(* IEC 61131-3 sources: plc-st-coding-agent/progress/evidence/f14_p1_20261111b/jobs/custom_minimax-m27 (part 2) *)

(* ---- self-hard-06.candidate_01.st ---- *)
FUNCTION_BLOCK FB
VAR_INPUT
    runRequest        : BOOL;
    pressure          : REAL;
    pressureValid     : BOOL;
    fuelFlow          : REAL;
    steamFlow         : REAL;
    outletCmd         : INT;
    outletFeedback    : INT;
    resetBtn          : BOOL;
END_VAR
VAR_OUTPUT
    tripLatched       : BOOL;
    fuelPermit        : BOOL;
    currentCauseMask  : WORD;
    latchedCauseMask  : WORD;
    diagnosticActive  : BOOL;
END_VAR
VAR
    stuckCount   : INT  := 0;      (* consecutive cycles for valve‑stuck detection *)
    prevResetBtn : BOOL := FALSE;   (* previous state of reset button *)
END_VAR

(* ------------------------------------------------------------------
   1. Valve‑stuck consecutive‑cycle detection
   ------------------------------------------------------------------ *)
IF runRequest AND pressureValid AND (pressure >= 4500.0)
   AND (outletCmd >= 50) AND (outletFeedback <= 10) THEN
    IF stuckCount < 3 THEN
        stuckCount := stuckCount + 1;
    END_IF;
ELSE
    stuckCount := 0;
END_IF;

(* ------------------------------------------------------------------
   2. Current cause mask (bits 0…3)
   ------------------------------------------------------------------ *)
IF NOT runRequest THEN
    currentCauseMask := 0;                     (* S5 *)

ELSIF NOT pressureValid THEN
    currentCauseMask := 1;                     (* bit0 – transmitter failure, S12 *)

ELSE
    (* pressureValid = TRUE *)
    IF pressure >= 4500.0 THEN
        (* Over‑pressure – evaluate bit1 (valve stuck) and bit2 (combustion excess) *)
        currentCauseMask := 0;

        IF stuckCount >= 3 THEN
            currentCauseMask := 2;             (* bit1 *)
        END_IF;

        IF (fuelFlow >= 4.0) AND (steamFlow <= 10.0) THEN
            currentCauseMask := currentCauseMask OR 4;  (* bit2 *)
        END_IF;

        (* If neither cause is identified, set bit3 (unlocated) *)
        IF currentCauseMask = 0 THEN
            currentCauseMask := 8;             (* bit3 *)
        END_IF;
    ELSE
        currentCauseMask := 0;                 (* S6 *)
    END_IF;
END_IF;

(* ------------------------------------------------------------------
   3. Trip condition
   ------------------------------------------------------------------ *)
(*  runRequest  AND ( pressureValid = FALSE  OR  pressure >= 4500.0 ) *)
tripLatched := tripLatched OR (runRequest AND (NOT pressureValid OR (pressure >= 4500.0)));

(* ------------------------------------------------------------------
   4. Reset on rising edge of reset button when conditions are met
   ------------------------------------------------------------------ *)
IF resetBtn AND NOT prevResetBtn AND NOT runRequest AND pressureValid AND (pressure <= 4200.0) THEN
    tripLatched := FALSE;
END_IF;
prevResetBtn := resetBtn;

(* ------------------------------------------------------------------
   5. Fuel permit
   ------------------------------------------------------------------ *)
fuelPermit := runRequest AND NOT tripLatched;   (* S3, N10‑S16 *)

(* ------------------------------------------------------------------
   6. Diagnostic active flag
   ------------------------------------------------------------------ *)
diagnosticActive := (currentCauseMask <> 0);    (* S7 *)

(* ------------------------------------------------------------------
   7. Accumulate cause mask while trip is latched
   ------------------------------------------------------------------ *)
IF tripLatched THEN
    latchedCauseMask := latchedCauseMask OR currentCauseMask;
ELSE
    latchedCauseMask := 0;                      (* N10‑S18 *)
END_IF;

END_FUNCTION_BLOCK

(* ---- self-medium-01.candidate_01.st ---- *)
TYPE ST_Recipe :
STRUCT
    recipeID   : INT;
    totalRatio : REAL;
    temperature: REAL;
END_STRUCT
END_TYPE

FUNCTION_BLOCK FB
VAR_INPUT
    recipe   : ARRAY[1..8] OF ST_Recipe;
    selSlot  : INT;
    loadCmd  : BOOL;
    running  : BOOL;
END_VAR
VAR_OUTPUT
    valid    : BOOL;
    loadedID : INT;
END_VAR
VAR
    prevLoadCmd  : BOOL := FALSE;
    prevRunning  : BOOL := FALSE;
    prevLoadedID : INT  := 0;
    prevValid    : BOOL := FALSE;
END_VAR
VAR_TEMP
    risingLoadCmd : BOOL;
    tmpRecipe     : ST_Recipe;
END_VAR

    // 检测 loadCmd 上升沿
    risingLoadCmd := loadCmd AND NOT prevLoadCmd;

    // 装载逻辑
    IF NOT running AND risingLoadCmd THEN
        // 槽位越界检查：必须先检查，不得访问数组外内存
        IF selSlot < 1 OR selSlot > 8 THEN
            valid   := FALSE;
            loadedID := 0;
        ELSE
            tmpRecipe := recipe[selSlot];
            // 槽位为空检查
            IF tmpRecipe.recipeID = 0 THEN
                valid   := FALSE;
                loadedID := 0;
            // 总配比越界检查 (99.0 <= totalRatio <= 101.0)
            ELSIF tmpRecipe.totalRatio < 99.0 OR tmpRecipe.totalRatio > 101.0 THEN
                valid   := FALSE;
                loadedID := 0;
            // 温度越界检查 (30.0 <= temperature <= 180.0)
            ELSIF tmpRecipe.temperature < 30.0 OR tmpRecipe.temperature > 180.0 THEN
                valid   := FALSE;
                loadedID := 0;
            ELSE
                valid    := TRUE;
                loadedID := tmpRecipe.recipeID;
            END_IF
        END_IF
    ELSE
        // 非装载周期：保持上一拍的值 (包括 running 状态)
        valid    := prevValid;
        loadedID := prevLoadedID;
    END_IF

    // 更新历史状态
    prevLoadCmd  := loadCmd;
    prevRunning  := running;
    prevLoadedID := loadedID;
    prevValid    := valid;

END_FUNCTION_BLOCK

(* ---- self-medium-02.candidate_01.st ---- *)
FUNCTION_BLOCK FB
VAR_INPUT
    enable    : BOOL;      (* 滤波使能，FALSE 时清空历史 *)
    rawValue  : REAL;      (* 本周期原始采样值 *)
END_VAR

VAR_OUTPUT
    filteredValue : REAL;  (* 滤波输出 *)
    windowFull    : BOOL;  (* 历史窗口已填满 8 个样本后置 TRUE *)
    sampleCount   : INT;   (* 当前窗口内有效样本数 0..8 *)
END_VAR

VAR
    buffer : ARRAY[0..7] OF REAL;  (* 8 点环形缓冲区 *)
    head   : INT := 0;             (* 下一写入位置 0..7 *)
    count  : INT := 0;             (* 有效样本数 0..8 *)
    full   : BOOL := FALSE;        (* 内部满窗标志 *)
END_VAR

VAR_TEMP
    sum : REAL;                    (* 临时累加和 *)
    idx : INT;                     (* 遍历索引 *)
    i   : INT;                     (* 循环计数器 *)
END_VAR

(*--------------------------------------------------------------------*)
(* 功能块主体                                                         *)
(*--------------------------------------------------------------------*)
IF enable THEN
    (* ----- 把新样本压入环形缓冲区 ----- *)
    buffer[head] := rawValue;                 (* 写入 *)
    head := (head + 1) MOD 8;                (* 头指针前移 *)
    IF count < 8 THEN
        count := count + 1;                  (* 样本计数 +1 *)
    END_IF
    full := (count = 8);                     (* 满窗标志 *)

ELSE
    (* ----- enable = FALSE：立即清零计数与满窗标志 ----- *)
    count := 0;
    full  := FALSE;
    (* head 保持不变，下一次 enable=TRUE 时会被覆盖 *)
END_IF

(* ----- 计算滤波输出（仅在有有效样本时） ----- *)
IF enable AND count > 0 THEN
    sum := 0.0;
    (*  oldest  = head - count (模 8) *)
    idx := (head - count + 8) MOD 8;
    FOR i := 0 TO count - 1 DO
        sum := sum + buffer[idx];
        idx := (idx + 1) MOD 8;
    END_FOR
    filteredValue := sum / INT_TO_REAL(count);   (* 算术平均 *)
END_IF
(* 当 enable=FALSE 时 filteredValue 保持不变 *)

(* ----- 输出信号 ----- *)
windowFull  := full;
sampleCount := count;

END_FUNCTION_BLOCK

(* ---- self-medium-03.candidate_01.st ---- *)
FUNCTION_BLOCK FB
VAR_INPUT
    openBtn    : BOOL;
    closeBtn   : BOOL;
    openLimit  : BOOL;
    closeLimit : BOOL;
    obstacle   : BOOL;
END_VAR

VAR_OUTPUT
    motorUp    : BOOL;
    motorDown  : BOOL;
    errorFlag  : BOOL;
END_VAR

VAR
    openBtnPrev    : BOOL := FALSE;
    closeBtnPrev   : BOOL := FALSE;
    combinedPrev   : BOOL := FALSE;
    prevMotorUp    : BOOL := FALSE;
    prevMotorDown  : BOOL := FALSE;
    prevErrorFlag  : BOOL := FALSE;
    state          : INT  := 0;   // 0=IDLE,1=OPENING,2=CLOSING,3=FAULT
END_VAR

(* Local auxiliary variables *)
VAR
    risingOpen     : BOOL;
    risingClose    : BOOL;
    risingCombined : BOOL;
    combinedNow    : BOOL;
    startOpen      : BOOL;
    startClose     : BOOL;
END_VAR

(* Detect combined button state *)
combinedNow    := openBtn AND closeBtn;

(* Detect rising edges *)
risingOpen     := openBtn   AND NOT openBtnPrev;
risingClose    := closeBtn  AND NOT closeBtnPrev;
risingCombined := combinedNow AND NOT combinedPrev;

(* Start conditions: new command from IDLE without fault and no obstacle *)
startOpen  := NOT prevMotorUp   AND NOT prevMotorDown   AND NOT prevErrorFlag
              AND risingOpen    AND NOT closeBtn AND NOT openLimit;

startClose := NOT prevMotorUp   AND NOT prevMotorDown   AND NOT prevErrorFlag
              AND risingClose   AND NOT openBtn  AND NOT closeLimit;

(* Motor commands according to S12 / S13 *)
motorUp   := NOT obstacle AND NOT openLimit
             AND (prevMotorUp OR startOpen);

motorDown := NOT obstacle AND NOT closeLimit
             AND (prevMotorDown OR startClose);

(* Error flag latch (S14) *)
errorFlag := obstacle OR (prevErrorFlag AND NOT risingCombined);

(* Optional state for external monitoring *)
IF errorFlag THEN
    state := 3;               (* FAULT *)
ELSIF motorUp THEN
    state := 1;               (* OPENING *)
ELSIF motorDown THEN
    state := 2;               (* CLOSING *)
ELSE
    state := 0;               (* IDLE *)
END_IF

(* Update previous values for next scan *)
openBtnPrev    := openBtn;
closeBtnPrev   := closeBtn;
combinedPrev   := combinedNow;
prevMotorUp    := motorUp;
prevMotorDown  := motorDown;
prevErrorFlag  := errorFlag;

END_FUNCTION_BLOCK

(* ---- self-medium-04.candidate_01.st ---- *)
FUNCTION_BLOCK FB
VAR_INPUT
    startBtn   : BOOL;
    resetBtn   : BOOL;
    doneSensor : BOOL;
    targetVol  : REAL;
    flowVol    : REAL;
END_VAR
VAR_OUTPUT
    valveOpen  : BOOL;
    fillsToday : INT;
END_VAR
VAR
    prev_startBtn   : BOOL := FALSE;
    prev_resetBtn   : BOOL := FALSE;
    prev_valveOpen  : BOOL := FALSE;
    currentFillVol  : REAL := 0.0;
    pendingConfirm  : BOOL := FALSE;
END_VAR

VAR
    risingStart : BOOL;
    risingReset : BOOL;
END_VAR

// 检测上升沿（基于上周期状态）
risingStart := startBtn AND NOT prev_startBtn;
risingReset := resetBtn  AND NOT prev_resetBtn;

// 复位处理（最高优先级）
IF risingReset THEN
    fillsToday      := 0;
    valveOpen       := FALSE;
    pendingConfirm  := FALSE;
    currentFillVol  := 0.0;
ELSE
    // 非复位时处理

    // 启动新瓶
    IF risingStart THEN
        // 取消上一瓶的待确认（如果有）
        pendingConfirm := FALSE;
        // 清零本瓶累计并开阀
        currentFillVol := 0.0;
        valveOpen      := TRUE;
    END_IF;

    // 灌装累计（阀开时）
    IF valveOpen THEN
        currentFillVol := currentFillVol + flowVol;
    END_IF;

    // 达标检测：累计达到或超过目标体积时立即关阀并设待确认
    IF valveOpen AND currentFillVol >= targetVol THEN
        valveOpen      := FALSE;
        pendingConfirm := TRUE;
    END_IF;

    // 确认检测：待确认且传感器为真时确认并计数
    IF pendingConfirm AND doneSensor THEN
        pendingConfirm := FALSE;
        IF fillsToday < 32767 THEN
            fillsToday := fillsToday + 1;
        END_IF;
    END_IF;
END_IF;

// 更新状态变量
prev_startBtn  := startBtn;
prev_resetBtn  := resetBtn;
prev_valveOpen := valveOpen;

END_FUNCTION_BLOCK

(* ---- self-medium-05.candidate_01.st ---- *)
(*====================================================================*)
(*  FUNCTION_BLOCK FB                                                *)
(*  Boiler steam‑quality accumulator with fuel consumption, revenue  *)
(*  and net‑profit.  All specifications from the problem statement   *)
(*  are implemented exactly.                                         *)
(*====================================================================*)
FUNCTION_BLOCK FB

VAR_INPUT
    enable       : BOOL;   (*计量使能*)
    resetBtn     : BOOL;   (*清零按钮 – 上升沿有效*)
    scanSeconds  : LREAL;  (*本周期时长 (s) , 合法 0 < dt ≤ 10*)
    steamFlow    : LREAL;  (*蒸汽流量 (kg/s) , 合法 0 … 90*)
    fuelFlow     : LREAL;  (*燃料流量 (kg/s) , 合法 0 … 6*)
    steamTemp    : LREAL;  (*蒸汽温度 (℃)*)
    steamPressure: LREAL;  (*蒸汽压力 (kPa)*)
END_VAR

VAR_OUTPUT
    qualified    : BOOL;   (*本周期蒸汽是否合格*)
    dataFault    : BOOL;   (*数据故障标志*)
    qualifiedTon : LREAL;  (*累计合格蒸汽产量 (t)*)
    fuelTon      : LREAL;  (*累计燃料消耗 (t)*)
    revenue      : LREAL;  (*累计收入 (元)*)
    cost         : LREAL;  (*累计成本 (元)*)
    netProfit    : LREAL;  (*累计净收益 (元) – 允许为负*)
END_VAR

VAR
    prevResetBtn : BOOL := FALSE;   (*上一拍的 resetBtn 状态，用于边沿检测*)
END_VAR

(*------------------------------------------------------------------*)
(*  临时变量，仅用于本周期内部计算                                   *)
VAR_TEMP
    risingReset : BOOL;            (*resetBtn 上升沿标志*)
END_VAR

(*------------------------------------------------------------------*)
(*  1) 上升沿检测                                                   *)
risingReset := resetBtn AND NOT prevResetBtn;

(*------------------------------------------------------------------*)
(*  2) 数据故障判据                                                 *)
dataFault := (scanSeconds <= 0.0) OR (scanSeconds > 10.0)
             OR (steamFlow < 0.0) OR (steamFlow > 90.0)
             OR (fuelFlow < 0.0)  OR (fuelFlow > 6.0);

(*------------------------------------------------------------------*)
(*  3) 合格判据 (闭区间)                                            *)
qualified := (steamTemp >= 447.0) AND (steamTemp <= 453.0)
             AND (steamPressure >= 3750.0) AND (steamPressure <= 3850.0);

(*------------------------------------------------------------------*)
(*  4) 累计逻辑 – 复位上升沿拥有最高优先级                           *)
IF risingReset THEN
    (* 复位拍：清零且本拍不再累计 *)
    qualifiedTon := 0.0;
    fuelTon      := 0.0;
ELSE
    (* 非复位拍：仅在 enable 且无故障时累计 *)
    IF enable AND NOT dataFault THEN
        (* 燃料消耗 – 只要使能且数据有效即累计 *)
        fuelTon := fuelTon + fuelFlow * scanSeconds / 1000.0;

        (* 合格蒸汽产量 – 额外要求本周期蒸汽合格 *)
        IF qualified THEN
            qualifiedTon := qualifiedTon + steamFlow * scanSeconds / 1000.0;
        END_IF;
    END_IF;
END_IF;

(*------------------------------------------------------------------*)
(*  5) 金额计算 (每拍都更新)                                        *)
revenue   := qualifiedTon * 280.0;   (*元 = t × 280*)
cost      := fuelTon      * 1500.0;  (*元 = t × 1500*)
netProfit := revenue - cost;

(*------------------------------------------------------------------*)
(*  6) 保持非负 (仅作防御性编程，实际运算已保证非负)                 *)
IF qualifiedTon < 0.0 THEN qualifiedTon := 0.0; END_IF;
IF fuelTon      < 0.0 THEN fuelTon      := 0.0; END_IF;
IF revenue      < 0.0 THEN revenue      := 0.0; END_IF;
IF cost         < 0.0 THEN cost         := 0.0; END_IF;

(*------------------------------------------------------------------*)
(*  7) 为下一拍准备边沿检测                                         *)
prevResetBtn := resetBtn;

END_FUNCTION_BLOCK

(* ---- public-easy-01.candidate_01.st ---- *)
PROGRAM AutomatedFillingLine
VAR
    (* Input variables *)
    bottleSensor           BOOL;
    cleaningConfirmButton  BOOL;
    fillingConfirmButton   BOOL;
    cappingConfirmButton   BOOL;
    packingConfirmButton   BOOL;
    finishedButton         BOOL;

    (* Output variables *)
    Pump_Motor             BOOL;
    Filling_Valve          BOOL;
    Capping_Machine        BOOL;
    Packing_Machine        BOOL;
    Completion_Light       BOOL;

    (* Internal state variable *)
    CurrentState           INT;
END_VAR

(* State definitions *)
CONST
    STATE_IDLE      := 0;
    STATE_CLEANING  := 1;
    STATE_FILLING   := 2;
    STATE_CAPPING   := 3;
    STATE_PACKING   := 4;
    STATE_COMPLETED := 5;
END_CONST

(* Initialize all outputs to FALSE *)
Pump_Motor       := FALSE;
Filling_Valve    := FALSE;
Capping_Machine  := FALSE;
Packing_Machine  := FALSE;
Completion_Light := FALSE;

(* State machine logic *)
CASE CurrentState OF

    STATE_IDLE:
        (* Reset all outputs *)
        Pump_Motor       := FALSE;
        Filling_Valve    := FALSE;
        Capping_Machine  := FALSE;
        Packing_Machine  := FALSE;
        Completion_Light := FALSE;

        (* Transition to CLEANING when bottle is detected *)
        IF bottleSensor THEN
            CurrentState := STATE_CLEANING;
        END_IF

    STATE_CLEANING:
        (* Activate cleaning pump *)
        Pump_Motor := TRUE;

        (* Transition to FILLING when cleaning is confirmed *)
        IF cleaningConfirmButton THEN
            CurrentState := STATE_FILLING;
        END_IF

    STATE_FILLING:
        (* Activate filling valve *)
        Filling_Valve := TRUE;

        (* Transition to CAPPING when filling is confirmed *)
        IF fillingConfirmButton THEN
            CurrentState := STATE_CAPPING;
        END_IF

    STATE_CAPPING:
        (* Activate capping machine *)
        Capping_Machine := TRUE;

        (* Transition to PACKING when capping is confirmed *)
        IF cappingConfirmButton THEN
            CurrentState := STATE_PACKING;
        END_IF

    STATE_PACKING:
        (* Activate packing machine *)
        Packing_Machine := TRUE;

        (* Transition to COMPLETED when packing is confirmed *)
        IF packingConfirmButton THEN
            CurrentState := STATE_COMPLETED;
        END_IF

    STATE_COMPLETED:
        (* Light up completion indicator *)
        Completion_Light := TRUE;

        (* Transition to IDLE when bottle is picked up *)
        IF finishedButton THEN
            CurrentState := STATE_IDLE;
        END_IF

END_CASE

(* ---- public-easy-01.candidate_02.st ---- *)
PROGRAM AutomatedFillingLine
VAR
    bottleSensor           BOOL;
    cleaningConfirmButton  BOOL;
    fillingConfirmButton   BOOL;
    cappingConfirmButton   BOOL;
    packingConfirmButton   BOOL;
    finishedButton         BOOL;

    Pump_Motor             BOOL;
    Filling_Valve          BOOL;
    Capping_Machine        BOOL;
    Packing_Machine        BOOL;
    Completion_Light       BOOL;

    CurrentState           INT := 0;
END_VAR

CASE CurrentState OF
    0:
        Pump_Motor       := FALSE;
        Filling_Valve    := FALSE;
        Capping_Machine  := FALSE;
        Packing_Machine  := FALSE;
        Completion_Light := FALSE;

        IF bottleSensor THEN
            CurrentState := 1;
        END_IF

    1:
        Pump_Motor := TRUE;

        IF cleaningConfirmButton THEN
            CurrentState := 2;
        END_IF

    2:
        Filling_Valve := TRUE;

        IF fillingConfirmButton THEN
            CurrentState := 3;
        END_IF

    3:
        Capping_Machine := TRUE;

        IF cappingConfirmButton THEN
            CurrentState := 4;
        END_IF

    4:
        Packing_Machine := TRUE;

        IF packingConfirmButton THEN
            CurrentState := 5;
        END_IF

    5:
        Completion_Light := TRUE;

        IF finishedButton THEN
            CurrentState := 0;
        END_IF

END_CASE

(* ---- public-easy-06.candidate_01.st ---- *)
PROGRAM AerationBlowerControl
VAR
    // Inputs
    DO_LOW                : BOOL;
    AERATION_E_STOP_NC    : BOOL;

    // Outputs
    BLOWER_RUN                    : BOOL;
    AERATION_BLOWER_CYCLE_COUNT   : UINT := 0;

    // Internal variables
    StartTimer        : TON;
    BlowerRunPrev     : BOOL := FALSE;
END_VAR

// ---------------------------------------------------------------------------
// Start Delay Logic
// ---------------------------------------------------------------------------
// Conditions for starting: DO is low AND emergency stop is inactive
IF DO_LOW AND AERATION_E_STOP_NC THEN
    // Start the 5-second delay timer
    StartTimer(IN := TRUE, PT := T#5S);

    // Enable blower only after timer completes
    IF StartTimer.Q THEN
        BLOWER_RUN := TRUE;
    ELSE
        BLOWER_RUN := FALSE;
    END_IF;
ELSE
    // Conditions not met - immediately disable blower
    BLOWER_RUN := FALSE;

    // Reset the start timer (timer IN = FALSE)
    StartTimer(IN := FALSE);
END_IF;

// ---------------------------------------------------------------------------
// Start Cycle Counting
// Detect FALSE-to-TRUE transition of BLOWER_RUN
// ---------------------------------------------------------------------------
IF BLOWER_RUN AND NOT BlowerRunPrev THEN
    AERATION_BLOWER_CYCLE_COUNT := AERATION_BLOWER_CYCLE_COUNT + 1;
END_IF;

// Store previous state for edge detection
BlowerRunPrev := BLOWER_RUN;

END_PROGRAM

(* ---- public-easy-06.candidate_02.st ---- *)
PROGRAM AerationBlowerControl
VAR_INPUT
    DO_LOW             : BOOL;
    AERATION_E_STOP_NC : BOOL;
END_VAR

VAR_OUTPUT
    BLOWER_RUN                    : BOOL;
    AERATION_BLOWER_CYCLE_COUNT   : UINT := 0;
END_VAR

VAR
    StartTimer    : TON;
    BlowerRunPrev : BOOL := FALSE;
END_VAR

// ---------------------------------------------------------------------------
// Start Delay Logic
// ---------------------------------------------------------------------------
// Conditions for starting: DO is low AND emergency stop is inactive
IF DO_LOW AND AERATION_E_STOP_NC THEN
    // Start the 5-second delay timer
    StartTimer(IN := TRUE, PT := T#5S);

    // Enable blower only after timer completes
    IF StartTimer.Q THEN
        BLOWER_RUN := TRUE;
    ELSE
        BLOWER_RUN := FALSE;
    END_IF;
ELSE
    // Conditions not met - immediately disable blower
    BLOWER_RUN := FALSE;

    // Reset the start timer
    StartTimer(IN := FALSE);
END_IF;

// ---------------------------------------------------------------------------
// Start Cycle Counting
// Detect FALSE-to-TRUE transition of BLOWER_RUN
// ---------------------------------------------------------------------------
IF BLOWER_RUN AND NOT BlowerRunPrev THEN
    AERATION_BLOWER_CYCLE_COUNT := AERATION_BLOWER_CYCLE_COUNT + 1;
END_IF;

// Store previous state for edge detection
BlowerRunPrev := BLOWER_RUN;

END_PROGRAM

(* ---- public-hard-01.candidate_02.st ---- *)
(* Material Proportioning Process Control *)
(* PLC Program in Structured Text (ST) *)

PROGRAM MaterialProportioning
VAR_INPUT
    estop           : BOOL;  (* Emergency Stop Signal: FALSE=Emergency stop triggered, TRUE=No emergency stop *)
    opeMode         : BOOL;  (* Operation Mode: FALSE=Manual, TRUE=Automatic *)
    valveAStart     : BOOL;  (* Valve A Start Button *)
    valveBStart     : BOOL;  (* Valve B Start Button *)
    valveCStart     : BOOL;  (* Valve C Start Button *)
    valveDStart     : BOOL;  (* Valve D Start Button *)
    mixMotorStart   : BOOL;  (* Mixing Motor Start Button *)
    autoStart       : BOOL;  (* Automatic Start Button *)
    processMode     : BOOL;  (* Process Mode *)
    levelSensor     : INT;   (* Liquid Level Sensor (unit cm) *)
    mixMotorComplete: BOOL;  (* Mixing Complete Signal *)
END_VAR

VAR_OUTPUT
    valveARun   : BOOL;  (* Valve A Run Command *)
    valveBRun   : BOOL;  (* Valve B Run Command *)
    valveCRun   : BOOL;  (* Valve C Run Command *)
    valveDRun   : BOOL;  (* Valve D Run Command *)
    mixMotorRun : BOOL;  (* Mixing Motor Run Command *)
END_VAR

VAR
    autoState         : INT := 0;
    prevAutoStart     : BOOL := FALSE;
    prevValveAStart   : BOOL := FALSE;
    prevValveBStart   : BOOL := FALSE;
    prevValveCStart   : BOOL := FALSE;
    prevValveDStart   : BOOL := FALSE;
    prevMixMotorStart : BOOL := FALSE;
END_VAR

(* Constants for state machine *)
CONST
    IDLE      := 0;
    FILL_A    := 1;
    FILL_B    := 2;
    FILL_C    := 3;
    MIXING    := 4;
    DISCHARGE := 5;
END_CONST

(* Emergency Stop - Highest Priority *)
IF NOT estop THEN
    valveARun    := FALSE;
    valveBRun    := FALSE;
    valveCRun    := FALSE;
    valveDRun    := FALSE;
    mixMotorRun  := FALSE;
    autoState    := IDLE;
    prevAutoStart := FALSE;
    prevValveAStart := FALSE;
    prevValveBStart := FALSE;
    prevValveCStart := FALSE;
    prevValveDStart := FALSE;
    prevMixMotorStart := FALSE;
    RETURN;
END_IF

(* Rising edge detection for manual mode buttons *)
IF valveAStart AND NOT prevValveAStart THEN
    valveARun := NOT valveARun;
END_IF

IF valveBStart AND NOT prevValveBStart THEN
    valveBRun := NOT valveBRun;
END_IF

IF valveCStart AND NOT prevValveCStart THEN
    valveCRun := NOT valveCRun;
END_IF

IF valveDStart AND NOT prevValveDStart THEN
    valveDRun := NOT valveDRun;
END_IF

IF mixMotorStart AND NOT prevMixMotorStart THEN
    mixMotorRun := NOT mixMotorRun;
END_IF

(* Update previous button states *)
prevValveAStart   := valveAStart;
prevValveBStart   := valveBStart;
prevValveCStart   := valveCStart;
prevValveDStart   := valveDStart;
prevMixMotorStart := mixMotorStart;

(* Mode Selection *)
IF opeMode THEN
    (* ========== AUTOMATIC MODE ========== *)

    (* Initialize manual control outputs to FALSE *)
    IF NOT prevValveAStart THEN valveARun := FALSE; END_IF
    IF NOT prevValveBStart THEN valveBRun := FALSE; END_IF
    IF NOT prevValveCStart THEN valveCRun := FALSE; END_IF
    IF NOT prevValveDStart THEN valveDRun := FALSE; END_IF
    IF NOT prevMixMotorStart THEN mixMotorRun := FALSE; END_IF

    (* Start automatic process on rising edge of autoStart *)
    IF autoStart AND NOT prevAutoStart THEN
        IF autoState = IDLE THEN
            autoState := FILL_A;
        END_IF
    END_IF
    prevAutoStart := autoStart;

    (* State Machine - Sequential Control *)
    IF autoState = FILL_A THEN
        valveARun := TRUE;
        (* When level reaches 50cm, close valve A and open valve B *)
        IF levelSensor >= 50 THEN
            autoState := FILL_B;
            valveARun := FALSE;
            valveBRun := TRUE;
        END_IF

    ELSIF autoState = FILL_B THEN
        valveBRun := TRUE;
        (* When level reaches 80cm, close valve B *)
        IF levelSensor >= 80 THEN
            valveBRun := FALSE;

            (* Check processMode for next step *)
            IF NOT processMode THEN
                (* processMode=false: Direct to mixing *)
                autoState   := MIXING;
                mixMotorRun := TRUE;
            ELSE
                (* processMode=true: Fill material C first *)
                autoState := FILL_C;
            END_IF
        END_IF

    ELSIF autoState = FILL_C THEN
        valveCRun := TRUE;
        (* When level reaches 100cm, close valve C and start mixing *)
        IF levelSensor >= 100 THEN
            autoState   := MIXING;
            valveCRun   := FALSE;
            mixMotorRun := TRUE;
        END_IF

    ELSIF autoState = MIXING THEN
        mixMotorRun := TRUE;
        (* When mixing complete signal received, stop motor *)
        IF mixMotorComplete THEN
            autoState   := DISCHARGE;
            mixMotorRun := FALSE;
        END_IF

    ELSIF autoState = DISCHARGE THEN
        valveDRun := TRUE;
        (* After discharge, return to idle - process complete *)
        autoState := IDLE;
    END_IF

ELSE
    (* ========== MANUAL MODE ========== *)
    (* Reset automatic state when switching to manual *)
    prevAutoStart := FALSE;
    autoState := IDLE;
END_IF

END_PROGRAM

(* ---- public-hard-03.candidate_01.st ---- *)
PROGRAM RecipeManagement
VAR
    // Inputs
    addRecipe        : BOOL;
    deleteRecipe     : BOOL;
    modifyRecipe     : BOOL;
    queryRecipe      : BOOL;
    recipeIn         : ST_Recipe;

    // Outputs
    recipeAdded          : BOOL;
    recipeDeleted        : BOOL;
    recipeModified       : BOOL;
    recipeQueryResult    : ST_Recipe;
    error            : BOOL;
    status           : WORD;

    // Input/Output
    recipe           : ARRAY[1..10] OF ST_Recipe;

    // Internal variables
    i               : INT;
    foundIndex      : INT;
    emptySlotIndex  : INT;
    hasDuplicate    : BOOL;
    hasEmptySlot    : BOOL;
    found           : BOOL;
END_VAR

//---------------------------------------------------------------------------
// Initialization - Clear outputs at the start of each cycle
//---------------------------------------------------------------------------
error            := FALSE;
status           := 16#0000;
recipeAdded      := FALSE;
recipeDeleted    := FALSE;
recipeModified   := FALSE;

// Initialize query result to empty recipe
recipeQueryResult.recipeID              := 0;
recipeQueryResult.ingredientType        := 0;
recipeQueryResult.ingredientRatio       := 0.0;
recipeQueryResult.productionTemperature := 0.0;

//---------------------------------------------------------------------------
// Query Recipe Operation
// Triggered when queryRecipe signal is TRUE
// Searches for recipe by recipeID and outputs result
//---------------------------------------------------------------------------
IF queryRecipe THEN
    found      := FALSE;
    foundIndex := 0;

    FOR i := 1 TO 10 DO
        IF recipe[i].recipeID = recipeIn.recipeID THEN
            found      := TRUE;
            foundIndex := i;
            EXIT; // Exit loop once found
        END_IF
    END_FOR

    IF found THEN
        // Recipe found - output to query result
        recipeQueryResult := recipe[foundIndex];
        error  := FALSE;
        status := 16#0000;
    ELSE
        // Recipe not found - error status 16#8001
        error  := TRUE;
        status := 16#8001;
    END_IF
END_IF

//---------------------------------------------------------------------------
// Add Recipe Operation
// Triggered when addRecipe signal is TRUE
// Adds new recipe to first available empty slot
//---------------------------------------------------------------------------
IF addRecipe THEN
    hasDuplicate   := FALSE;
    hasEmptySlot   := FALSE;
    emptySlotIndex := 0;
    found          := FALSE;
    foundIndex     := 0;

    // Step 1: Check for duplicate recipeID
    FOR i := 1 TO 10 DO
        IF recipe[i].recipeID = recipeIn.recipeID THEN
            hasDuplicate := TRUE;
            found        := TRUE;
            EXIT;
        END_IF
    END_FOR

    IF hasDuplicate THEN
        // Duplicate recipeID found - error status 16#8002
        error  := TRUE;
        status := 16#8002;
    ELSE
        // Step 2: Find first empty slot (smallest index)
        FOR i := 1 TO 10 DO
            IF recipe[i].recipeID = 0 THEN
                hasEmptySlot   := TRUE;
                emptySlotIndex := i;
                EXIT;
            END_IF
        END_FOR

        IF NOT hasEmptySlot THEN
            // No empty slot available - error status 16#8003
            error  := TRUE;
            status := 16#8003;
        ELSE
            // Step 3: Store recipe in empty slot with smallest index
            recipe[emptySlotIndex] := recipeIn;
            recipeAdded            := TRUE;
            error                  := FALSE;
            status                 := 16#0000;
        END_IF
    END_IF
END_IF

//---------------------------------------------------------------------------
// Delete Recipe Operation
// Triggered when deleteRecipe signal is TRUE
// Sets recipeID to 0 (marks slot as empty)
//---------------------------------------------------------------------------
IF deleteRecipe THEN
    found      := FALSE;
    foundIndex := 0;

    // Search for recipe by recipeID
    FOR i := 1 TO 10 DO
        IF recipe[i].recipeID = recipeIn.recipeID THEN
            found      := TRUE;
            foundIndex := i;
            EXIT;
        END_IF
    END_FOR

    IF found THEN
        // Recipe found - delete by setting recipeID to 0
        recipe[foundIndex].recipeID              := 0;
        recipe[foundIndex].ingredientType        := 0;
        recipe[foundIndex].ingredientRatio       := 0.0;
        recipe[foundIndex].productionTemperature := 0.0;
        recipeDeleted                            := TRUE;
        error                                    := FALSE;
        status                                   := 16#0000;
    ELSE
        // Recipe not found - error status 16#8004
        error  := TRUE;
        status := 16#8004;
    END_IF
END_IF

//---------------------------------------------------------------------------
// Modify Recipe Operation
// Triggered when modifyRecipe signal is TRUE
// Replaces existing recipe with input recipe
//---------------------------------------------------------------------------
IF modifyRecipe THEN
    found      := FALSE;
    foundIndex := 0;

    // Search for recipe by recipeID
    FOR i := 1 TO 10 DO
        IF recipe[i].recipeID = recipeIn.recipeID THEN
            found      := TRUE;
            foundIndex := i;
            EXIT;
        END_IF
    END_FOR

    IF found THEN
        // Recipe found - replace with input recipe
        recipe[foundIndex] := recipeIn;
        recipeModified     := TRUE;
        error              := FALSE;
        status             := 16#0000;
    ELSE
        // Recipe not found - error status 16#8005
        error  := TRUE;
        status := 16#8005;
    END_IF
END_IF

END_PROGRAM

(* ---- public-hard-06.candidate_01.st ---- *)
(*----------------------------------------------------------------------------------
  Production Line Controller – Hard Version
  Mode 0 = Manual, Mode 1 = Automatic
  Automatic sequence: Feed → Wash → Weigh → Fire → Output
  Manual mode: forward / reverse with interlock
----------------------------------------------------------------------------------*)

(*----------- Type definitions ----------------------------------------------------*)
TYPE E_State :
(
    IDLE             := 0,
    MOVING_TO_WASH   := 1,
    AT_WASH          := 2,
    MOVING_TO_WEIGH  := 3,
    AT_WEIGH         := 4,
    MOVING_TO_FIRING := 5,
    AT_FIRING        := 6,
    MOVING_TO_OUTPUT := 7,
    AT_OUTPUT        := 8,
    REJECT           := 9
);
END_TYPE

(*----------- Program declaration -------------------------------------------------*)
PROGRAM ProductionControl
VAR_INPUT
    Mode            : BOOL;          (* 0 = Manual, 1 = Automatic *)
    ForwardButton   : BOOL;          (* Manual forward command *)
    ReverseButton   : BOOL;          (* Manual reverse command *)
    SensorFeed      : BOOL;          (* Material at loading station *)
    SensorWash      : BOOL;          (* Material at cleaning station *)
    SensorWeight    : BOOL;          (* Material at weighing station *)
    SensorFiring    : BOOL;          (* Product at firing station *)
    SensorOutput    : BOOL;          (* Product at finished‑product station *)
    washComplete    : BOOL;          (* Cleaning finished *)
    weightComplete  : BOOL;          (* Weighing finished *)
    weight          : REAL;          (* Measured weight *)
    firingComplete  : BOOL;          (* Firing finished *)
END_VAR

VAR_OUTPUT
    MotorForward    : BOOL;          (* Motor forward rotation *)
    MotorReverse    : BOOL;          (* Motor reverse rotation *)
    kick            : BOOL;          (* Rejection command *)
    CompletionLight : BOOL;          (* Product ready light *)
    firingTemp      : REAL;          (* Calculated firing temperature *)
END_VAR

(*----------- Internal variables -------------------------------------------------*)
VAR
    curState        : E_State := IDLE;   (* Current automatic state *)

    (* Edge detection memories *)
    lastSensorFeed    : BOOL := FALSE;
    lastSensorWash    : BOOL := FALSE;
    lastSensorWeight  : BOOL := FALSE;
    lastSensorFiring  : BOOL := FALSE;
    lastSensorOutput  : BOOL := FALSE;
    lastWashComplete  : BOOL := FALSE;
    lastWeightComplete: BOOL := FALSE;
    lastFiringComplete: BOOL := FALSE;

    (* Edge flags *)
    sensorFeedRising    : BOOL;
    sensorWashRising    : BOOL;
    sensorWeightRising  : BOOL;
    sensorFiringRising  : BOOL;
    sensorOutputRising  : BOOL;
    sensorOutputFalling : BOOL;
    washCompleteRising  : BOOL;
    weightCompleteRising: BOOL;
    firingCompleteRising: BOOL;

    (* One‑shot flags for completion signals *)
    washProcessed   : BOOL := FALSE;
    weightProcessed : BOOL := FALSE;
    firingProcessed : BOOL := FALSE;
END_VAR

(*----------- Edge detection ----------------------------------------------------*)
sensorFeedRising     := SensorFeed     AND NOT lastSensorFeed;
sensorWashRising     := SensorWash     AND NOT lastSensorWash;
sensorWeightRising   := SensorWeight   AND NOT lastSensorWeight;
sensorFiringRising   := SensorFiring   AND NOT lastSensorFiring;
sensorOutputRising   := SensorOutput   AND NOT lastSensorOutput;
sensorOutputFalling  := NOT SensorOutput AND lastSensorOutput;

washCompleteRising   := washComplete   AND NOT lastWashComplete;
weightCompleteRising := weightComplete AND NOT lastWeightComplete;
firingCompleteRising := firingComplete AND NOT lastFiringComplete;

(* Update memories *)
lastSensorFeed    := SensorFeed;
lastSensorWash    := SensorWash;
lastSensorWeight  := SensorWeight;
lastSensorFiring  := SensorFiring;
lastSensorOutput  := SensorOutput;
lastWashComplete  := washComplete;
lastWeightComplete:= weightComplete;
lastFiringComplete:= firingComplete;

(*----------- Mode handling ------------------------------------------------------*)
IF Mode = FALSE THEN                (* Manual Mode *)
    (* Reset automatic control outputs *)
    MotorForward    := FALSE;
    MotorReverse    := FALSE;
    kick            := FALSE;
    CompletionLight := FALSE;
    firingTemp      := 0.0;
    curState        := IDLE;
    washProcessed   := FALSE;
    weightProcessed := FALSE;
    firingProcessed := FALSE;

    (* Interlocked forward / reverse *)
    IF ForwardButton AND NOT ReverseButton THEN
        MotorForward := TRUE;
    ELSE
        MotorForward := FALSE;
    END_IF

    IF ReverseButton AND NOT ForwardButton THEN
        MotorReverse := TRUE;
    ELSE
        MotorReverse := FALSE;
    END_IF

ELSE                                 (* Automatic Mode *)
    MotorReverse := FALSE;          (* Reverse never used in auto *)

    CASE curState OF

        (*--------------------------------------------------------------
         IDLE – waiting for a new material at the loading station
        --------------------------------------------------------------*)
        IDLE:
            IF sensorFeedRising THEN
                curState     := MOVING_TO_WASH;
                MotorForward := TRUE;
            ELSE
                MotorForward    := FALSE;
                kick            := FALSE;
                CompletionLight := FALSE;
                firingTemp      := 0.0;
            END_IF

        (*--------------------------------------------------------------
         MOVING_TO_WASH – motor conveys material to cleaning station
        --------------------------------------------------------------*)
        MOVING_TO_WASH:
            IF sensorWashRising THEN
                MotorForward := FALSE;
                curState     := AT_WASH;
                washProcessed := FALSE;
            END_IF

        (*--------------------------------------------------------------
         AT_WASH – cleaning in progress, waiting for washComplete
        --------------------------------------------------------------*)
        AT_WASH:
            IF washCompleteRising AND NOT washProcessed THEN
                MotorForward := TRUE;
                curState      := MOVING_TO_WEIGH;
                washProcessed := TRUE;
            END_IF

        (*--------------------------------------------------------------
         MOVING_TO_WEIGH – material moves to weighing station
        --------------------------------------------------------------*)
        MOVING_TO_WEIGH:
            IF sensorWeightRising THEN
                MotorForward   := FALSE;
                curState       := AT_WEIGH;
                weightProcessed := FALSE;
            END_IF

        (*--------------------------------------------------------------
         AT_WEIGH – weight measurement, quality check and temperature calc.
        --------------------------------------------------------------*)
        AT_WEIGH:
            IF weightCompleteRising AND NOT weightProcessed THEN
                weightProcessed := TRUE;
                IF weight >= 100.0 AND weight <= 200.0 THEN
                    (* Qualified – compute firing temperature *)
                    firingTemp  := 500.0 + ((weight - 100.0) / 100.0) * 50.0;
                    MotorForward := TRUE;
                    curState     := MOVING_TO_FIRING;
                ELSE
                    (* Unqualified – reject *)
                    kick         := TRUE;
                    MotorForward := FALSE;
                    curState     := REJECT;
                END_IF
            END_IF

        (*--------------------------------------------------------------
         MOVING_TO_FIRING – material moves to firing station
        --------------------------------------------------------------*)
        MOVING_TO_FIRING:
            IF sensorFiringRising THEN
                MotorForward   := FALSE;
                curState       := AT_FIRING;
                firingProcessed := FALSE;
            END_IF

        (*--------------------------------------------------------------
         AT_FIRING – firing in progress, waiting for firingComplete
        --------------------------------------------------------------*)
        AT_FIRING:
            IF firingCompleteRising AND NOT firingProcessed THEN
                MotorForward   := TRUE;
                curState        := MOVING_TO_OUTPUT;
                firingProcessed := TRUE;
            END_IF

        (*--------------------------------------------------------------
         MOVING_TO_OUTPUT – product moves to finished‑product station
        --------------------------------------------------------------*)
        MOVING_TO_OUTPUT:
            IF sensorOutputRising THEN
                MotorForward    := FALSE;
                CompletionLight := TRUE;
                curState        := AT_OUTPUT;
            END_IF

        (*--------------------------------------------------------------
         AT_OUTPUT – product waiting to be taken away
        --------------------------------------------------------------*)
        AT_OUTPUT:
            CompletionLight := SensorOutput;   (* Light on while product present *)
            IF sensorOutputFalling THEN
                CompletionLight := FALSE;
                curState        := IDLE;
                firingTemp      := 0.0;
                kick            := FALSE;
            END_IF

        (*--------------------------------------------------------------
         REJECT – unqualified material at weighing station
        --------------------------------------------------------------*)
        REJECT:
            kick         := TRUE;
            MotorForward := FALSE;
            (* Assume the material is removed manually; when weight sensor clears → reset *)
            IF NOT SensorWeight THEN
                kick     := FALSE;
                curState := IDLE;
            END_IF

    END_CASE
END_IF

END_PROGRAM

(* ---- public-medium-07.candidate_01.st ---- *)
(* -------------------------------------------------------------
   Office HVAC Multi‑mode Energy‑Saving Control
   -------------------------------------------------------------
   Inputs
     OCCUPANCY_DETECTED   – TRUE when occupancy is detected
     ENERGY_SAVING_MODE   – TRUE → energy‑saving, FALSE → standard
     HVAC_MODE_SELECTOR   – 0 = Auto, 1 = Comfort, 2 = Economy, 3 = Night
   Outputs
     SUPPLY_FAN_RUN       – Supply‑fan run enable (BOOL)
     TEMP_SETPOINT_ADJUST – Temperature‑setpoint adjustment in °C (INT)
   -------------------------------------------------------------
   Behaviour
     • 30 s on‑delay for the fan when occupied and NOT in Night mode.
       The fan is stopped immediately and the timer is reset when
       occupancy is lost or Night mode is entered.
     • Temperature‑setpoint adjustment follows the table:
       Mode   | Occupied | Unoccupied (standard) | Unoccupied (energy‑saving)
       -------|----------|-----------------------|----------------------------
       Auto   |   0 °C   |        +2 °C          |            +3 °C
       Comfort|   0 °C   |        +1 °C          |            +1 °C
       Economy|   0 °C   |        +4 °C          |            +4 °C
       Night  |   +4 °C  |        +4 °C          |            +4 °C
       (Energy‑saving flag influences only Auto mode.)
     • Outputs are initialised to OFF / 0 at power‑up and are updated
       every scan from the current inputs.
   ------------------------------------------------------------- *)

PROGRAM HVAC_Control
   VAR_INPUT
      OCCUPANCY_DETECTED   : BOOL;
      ENERGY_SAVING_MODE   : BOOL;
      HVAC_MODE_SELECTOR   : INT;
   END_VAR

   VAR_OUTPUT
      SUPPLY_FAN_RUN       : BOOL := FALSE;   (* OFF at power‑up *)
      TEMP_SETPOINT_ADJUST : INT  := 0;       (* zero at power‑up *)
   END_VAR

   VAR
      FanTimer      : TON;                    (* 30‑second on‑delay *)
      FanStartCond  : BOOL;                   (* condition to start the timer *)
   END_VAR

   (* ---------------------------------------------------------
      Fan start condition: occupied AND NOT Night mode
      --------------------------------------------------------- *)
   FanStartCond := OCCUPANCY_DETECTED AND (HVAC_MODE_SELECTOR <> 3);

   (* ---------------------------------------------------------
      30‑second ON‑delay timer
      The timer resets automatically when FanStartCond becomes FALSE,
      fulfilling the “reset timing if occupancy is lost or Night mode
      is selected” requirement.
      --------------------------------------------------------- *)
   FanTimer(IN := FanStartCond, PT := T#30s);
   SUPPLY_FAN_RUN := FanTimer.Q;

   (* ---------------------------------------------------------
      Temperature‑setpoint adjustment according to mode,
      occupancy and energy‑saving selection.
      --------------------------------------------------------- *)
   CASE HVAC_MODE_SELECTOR OF
      0 : (* Auto *)
         IF OCCUPANCY_DETECTED THEN
            TEMP_SETPOINT_ADJUST := 0;
         ELSE
            IF ENERGY_SAVING_MODE THEN
               TEMP_SETPOINT_ADJUST := 3;   (* +3 °C when energy‑saving *)
            ELSE
               TEMP_SETPOINT_ADJUST := 2;   (* +2 °C in standard mode *)
            END_IF;
         END_IF;

      1 : (* Comfort *)
         IF OCCUPANCY_DETECTED THEN
            TEMP_SETPOINT_ADJUST := 0;
         ELSE
            TEMP_SETPOINT_ADJUST := 1;
         END_IF;

      2 : (* Economy *)
         IF OCCUPANCY_DETECTED THEN
            TEMP_SETPOINT_ADJUST := 0;
         ELSE
            TEMP_SETPOINT_ADJUST := 4;
         END_IF;

      3 : (* Night *)
         TEMP_SETPOINT_ADJUST := 4;

   END_CASE;

END_PROGRAM
